(* IEC 61131-3 sources: llm-plc-st-eval/data/processed/gpt-4o/B3/few_shot, 3 files *)

(* ---- ejec_1.st ---- *)
FUNCTION_BLOCK FB_Contador
VAR_INPUT
    sensorPieza : BOOL; (* Sensor fotoeléctrico para detectar piezas *)
    btnReset : BOOL;    (* Botón para resetear el contador *)
END_VAR
VAR_OUTPUT
    loteListo : BOOL;   (* Indica si el lote está completo *)
    cuenta : INT;       (* Cuenta de piezas detectadas *)
END_VAR
VAR
    sensorPiezaAnt : BOOL; (* Estado anterior del sensor de pieza *)
END_VAR

(* Inicialización de variables *)
IF btnReset THEN
    cuenta := 0;
    loteListo := FALSE;
ELSE
    (* Detectar transición de FALSE a TRUE en el sensor de pieza *)
    IF (sensorPieza AND NOT sensorPiezaAnt) THEN
        cuenta := cuenta + 1;
    END_IF;

    (* Verificar si se ha alcanzado el conteo de 12 piezas *)
    IF cuenta >= 12 THEN
        loteListo := TRUE;
    ELSE
        loteListo := FALSE;
    END_IF;
END_IF;

(* Actualizar el estado anterior del sensor de pieza *)
sensorPiezaAnt := sensorPieza;
END_FUNCTION_BLOCK

(* ---- ejec_2.st ---- *)
FUNCTION_BLOCK FB_Contador
VAR_INPUT
    sensorPieza : BOOL; (* Sensor fotoeléctrico para detección de piezas *)
    btnReset : BOOL;    (* Botón para reiniciar el contador *)
END_VAR
VAR_OUTPUT
    loteListo : BOOL;   (* Indica si el lote está completo *)
    cuenta : INT;       (* Cuenta de piezas detectadas *)
END_VAR
VAR
    sensorPiezaAnt : BOOL; (* Estado anterior del sensor de pieza *)
END_VAR

(* Inicialización de variables *)
IF btnReset THEN
    cuenta := 0;
    loteListo := FALSE;
ELSE
    (* Detecta la transición de FALSE a TRUE del sensor de pieza *)
    IF (sensorPieza AND NOT sensorPiezaAnt) THEN
        cuenta := cuenta + 1;
    END_IF;

    (* Verifica si se ha alcanzado el conteo de 12 piezas *)
    IF cuenta >= 12 THEN
        loteListo := TRUE;
    ELSE
        loteListo := FALSE;
    END_IF;
END_IF;

(* Actualiza el estado anterior del sensor de pieza *)
sensorPiezaAnt := sensorPieza;
END_FUNCTION_BLOCK

(* ---- ejec_3.st ---- *)
FUNCTION_BLOCK FB_Contador
VAR_INPUT
    sensorPieza : BOOL; (* Sensor fotoeléctrico para detección de piezas *)
    btnReset : BOOL;    (* Botón para resetear el contador *)
END_VAR
VAR_OUTPUT
    loteListo : BOOL;   (* Indica si el lote está completo *)
    cuenta : INT;       (* Contador de piezas *)
END_VAR
VAR
    sensorPiezaAnt : BOOL; (* Estado anterior del sensor de pieza *)
END_VAR

(* Detectar flanco ascendente del sensor de pieza *)
IF NOT sensorPiezaAnt AND sensorPieza THEN
    cuenta := cuenta + 1; (* Incrementar cuenta en flanco ascendente *)
END_IF

(* Resetear el contador y la salida de lote completo *)
IF btnReset THEN
    cuenta := 0;
    loteListo := FALSE;
END_IF

(* Verificar si el lote está completo *)
IF cuenta >= 12 THEN
    loteListo := TRUE;
ELSE
    loteListo := FALSE;
END_IF

(* Actualizar el estado anterior del sensor de pieza *)
sensorPiezaAnt := sensorPieza;

END_FUNCTION_BLOCK
